// TIA Portal project "Project3" (V13)

(* hardware
DEVICE "S7-1200 station_1"  S7-1200 Station
   slot 0: "Rack_0"  Rack  V1.0
   slot 1: "PLC_1"  CPU 1212C AC/DC/Rly  6ES7 212-1BE40-0XB0  V4.1
DEVICE "GSD device_1"  GSD.Device.PN
   slot 0: "Rack"  Rail  V1.0
   slot 0: "AL1100"  AL1100
   slot 1: "4 Ports_1"  AL1100
DEVICE "HMI_2"  KTP400 Basic PN
   slot 0: "HMI"  HMI  6AV2 123-2DB03-0AX0  13.0.0.0
   slot 1: "HMI_RT_2"  KTP400 Basic PN  6AV2 123-2DB03-0AX0  13.0.0.0
   slot 5: "HMI_2.IE_CP_1"  PROFINET Interface
      slot 1: "PROFINET Interface_1"  PROFINET Interface
         slot 1: "Port_1"  Port
*)

// ===== PLC "PLC_1"  CPU 1212C AC/DC/Rly =====

VAR_GLOBAL   // PLC tag table "Default tag table"
   "Tag_1" AT %Q0.0 : Bool;
   "Tag_2" AT %M0.0 : Bool;
   "System_Byte" AT %MB1 : Byte;
   "FirstScan" AT %M1.0 : Bool;
   "DiagStatusUpdate" AT %M1.1 : Bool;
   "AlwaysTRUE" AT %M1.2 : Bool;
   "AlwaysFALSE" AT %M1.3 : Bool;
   "Clock_Byte" AT %MB0 : Byte;
   "Clock_5Hz" AT %M0.1 : Bool;
   "Clock_2.5Hz" AT %M0.2 : Bool;
   "Clock_2Hz" AT %M0.3 : Bool;
   "Clock_1.25Hz" AT %M0.4 : Bool;
   "Clock_1Hz" AT %M0.5 : Bool;
   "Clock_0.625Hz" AT %M0.6 : Bool;
   "Clock_0.5Hz" AT %M0.7 : Bool;
   "Tag_3" AT %M10.0 : Bool;
END_VAR

VAR_GLOBAL   // PLC tag table "RFID"
   "i_command_value" AT %IB90 : Byte;
   "i_command_ack" AT %I91.0 : Bool;
   "i_command_end" AT %I91.1 : Bool;
   "i_tag_present" AT %I91.2 : Bool;
   "i_antenna_deactivated" AT %I91.3 : Bool;
   "i_read_value_0" AT %IW92 : Int;
   "i_read_value_1" AT %IW94 : Int;
   "i_read_value_2" AT %IW96 : Int;
   "i_read_value_3" AT %IW98 : Int;
   "q_command_value" AT %QB84 : Byte;
   "q_start_r/w" AT %Q85.0 : Bool;
   "q_antenna_deactivate" AT %Q85.3 : Bool;
   "q_write_value_0" AT %QW86 : Int;
   "q_write_value_1" AT %QW88 : Int;
   "q_write_value_2" AT %QW90 : Int;
   "q_write_value_3" AT %QW92 : Int;
END_VAR

TYPE "RFID_IOLink"
   STRUCT
      Input : Struct
      END_STRUCT;
      Output : Struct
      END_STRUCT;
   END_STRUCT;
END_TYPE

DATA_BLOCK "test"   // DB2
{ S7_Optimized_Access := 'FALSE' }
VERSION : 0.1
   VAR
      demo : Bool;
      data : Int;
   END_VAR
BEGIN
END_DATA_BLOCK

DATA_BLOCK "Logic_DB"   // DB4
{ S7_Optimized_Access := 'FALSE' }
VERSION : 0.1
// stored: InstanceOfName Logic
"Logic"
BEGIN
END_DATA_BLOCK

// folder: RFID

DATA_BLOCK "RFIDData"   // DB1
{ S7_Optimized_Access := 'FALSE' }
VERSION : 0.1
   VAR
      RFID : "RFID_IOLink";
   END_VAR
BEGIN
END_DATA_BLOCK

DATA_BLOCK "Logic DB"   // DB3
{ S7_Optimized_Access := 'FALSE' }
VERSION : 0.1
   VAR
      TimeParameters : Struct
      END_STRUCT;
      BufferControl : Struct
      END_STRUCT;
      Error : Struct
      END_STRUCT;
   END_VAR
BEGIN
END_DATA_BLOCK

DATA_BLOCK "BufferData_DB"   // DB5
{ S7_Optimized_Access := 'FALSE' }
VERSION : 0.1
// stored: InstanceOfName BufferData
"BufferData"
BEGIN
END_DATA_BLOCK

// folder: (top level)

ORGANIZATION_BLOCK "Main"   // OB1, LAD, ProgramCycle
TITLE = "Main Program Sweep (Cycle)"
{ S7_Optimized_Access := 'FALSE' }
VERSION : 0.1
BEGIN

REGION Network 1: Read values from RFID
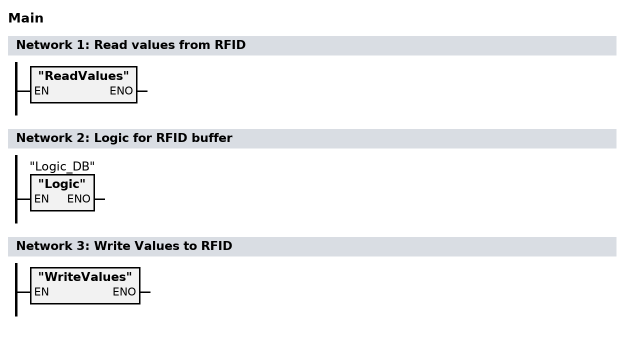
   RUNG wire#powerrail
      "ReadValues"()
   END_RUNG
   // the same network as SCL:
   "ReadValues"();
END_REGION

REGION Network 2: Logic for RFID buffer
   RUNG wire#powerrail
      "Logic_DB"()
   END_RUNG
   // the same network as SCL:
   "Logic_DB"();   // "Logic"
END_REGION

REGION Network 3: Write Values to RFID
   RUNG wire#powerrail
      "WriteValues"()
   END_RUNG
   // the same network as SCL:
   "WriteValues"();
END_REGION
END_ORGANIZATION_BLOCK

// folder: RFID

FUNCTION_BLOCK "Logic"   // FB1, FBD
{ S7_Optimized_Access := 'FALSE' }
VERSION : 0.1
BEGIN

REGION Network 1: Log of tags with timestamp
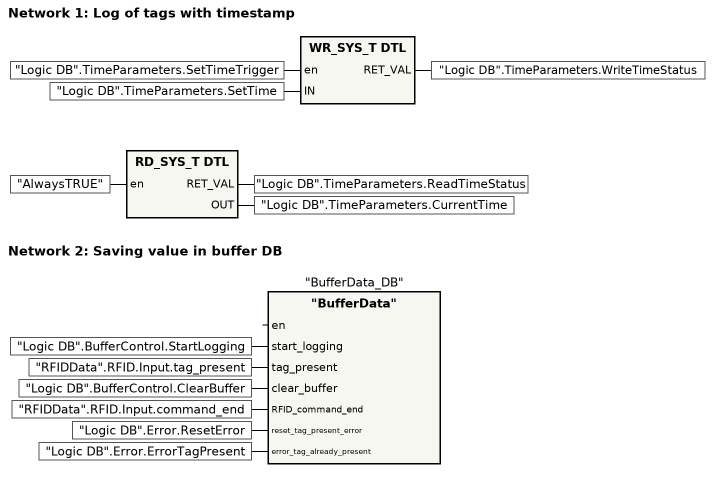
   IF "Logic DB".TimeParameters.SetTimeTrigger THEN
       "Logic DB".TimeParameters.WriteTimeStatus := WR_SYS_T(IN := "Logic DB".TimeParameters.SetTime);
   END_IF;
   IF "AlwaysTRUE" THEN
       "Logic DB".TimeParameters.ReadTimeStatus := RD_SYS_T(OUT => "Logic DB".TimeParameters.CurrentTime);
   END_IF;
END_REGION

REGION Network 2: Saving value in buffer DB
   "BufferData_DB"(start_logging := "Logic DB".BufferControl.StartLogging,   // "BufferData"
                   tag_present := "RFIDData".RFID.Input.tag_present,
                   clear_buffer := "Logic DB".BufferControl.ClearBuffer,
                   RFID_command_end := "RFIDData".RFID.Input.command_end,
                   reset_tag_present_error := "Logic DB".Error.ResetError,
                   error_tag_already_present := "Logic DB".Error.ErrorTagPresent);
END_REGION
END_FUNCTION_BLOCK

FUNCTION_BLOCK "BufferData"   // FB2, SCL
{ S7_Optimized_Access := 'FALSE' }
VERSION : 0.1
BEGIN
   //Generating rising edge bit for RFID 'End' status
   #command_end_flag:= #RFID_command_end AND NOT #M_command_end_flag;
   #M_command_end_flag := #RFID_command_end;

   //Check tag validity i.e. Tag should not be = 0 and not already registered
   IF (#start_logging AND NOT #error_tag_already_present) THEN
       IF (#command_end_flag) AND ("RFIDData".RFID.Input.read_values[0] <> 0) THEN 
           FOR #c := 0 TO 5 DO
               IF ("Logic DB".BufferControl.Job[#c].RFID = "RFIDData".RFID.Input.read_values[0]) THEN
                   #error_tag_already_present := true;
                   GOTO x2;
               END_IF;
           END_FOR;
   //IF RFID tag is not registered --> Registering the tag information in the next available slot
           FOR #d := 0 TO 5 DO
               IF (#command_end_flag) AND ("Logic DB".BufferControl.Job[#d].RFID = 0) AND NOT #error_tag_already_present THEN
                   "Logic DB".BufferControl.Job[#d].Job_ID := #d +1;
                   "Logic DB".BufferControl.Job[#d].RFID := "RFIDData".RFID.Input.read_values[0];
                   "Logic DB".BufferControl.Job[#d].ProcessTime :="Logic DB".TimeParameters.CurrentTime ;
                   GOTO x2;
               END_IF;
           END_FOR;
       x2: ;
      END_IF;
   END_IF;

   //Clear log button
   IF #clear_buffer THEN
       FOR #i := 0 TO 5 DO
           "Logic DB".BufferControl.Job[#i].ProcessTime := "Logic DB".TimeParameters.ResetTime;
           "Logic DB".BufferControl.Job[#i].RFID := 0;
           "Logic DB".BufferControl.Job[#i].Job_ID := 0;
       END_FOR;

   END_IF;

   IF (#reset_tag_present_error) THEN
       #error_tag_already_present := false;
   END_IF;
END_FUNCTION_BLOCK

FUNCTION "ReadValues" : Void   // FC1, SCL
{ S7_Optimized_Access := 'FALSE' }
VERSION : 0.1
BEGIN
   //Reading value from RFID
   "RFIDData".RFID.Input.command_ack:="i_command_ack";
   "RFIDData".RFID.Input.command_value:="i_command_value";
   "RFIDData".RFID.Input.command_end:="i_command_end";
   "RFIDData".RFID.Input.tag_present:="i_tag_present";
   "RFIDData".RFID.Input.Antenna_deactivated:="i_antenna_deactivated";
   "RFIDData".RFID.Input.read_values[0]:="i_read_value_0";
   "RFIDData".RFID.Input.read_values[1]:="i_read_value_1";
   "RFIDData".RFID.Input.read_values[2]:="i_read_value_2";
   "RFIDData".RFID.Input.read_values[3]:="i_read_value_3";
END_FUNCTION

FUNCTION "WriteValues" : Void   // FC2, SCL
{ S7_Optimized_Access := 'FALSE' }
VERSION : 0.1
BEGIN
   //Writing values to RFID
   "q_command_value" := "RFIDData".RFID.Output.command_value;
   "q_start_r/w" := "RFIDData".RFID.Output."Start_r/w";
   "q_antenna_deactivate" := "RFIDData".RFID.Output.Deactivate_antenna;
   "q_write_value_0" := "RFIDData".RFID.Output.write_values[0];
   "q_write_value_1" := "RFIDData".RFID.Output.write_values[1];
   "q_write_value_2" := "RFIDData".RFID.Output.write_values[2];
   "q_write_value_3" := "RFIDData".RFID.Output.write_values[3];
END_FUNCTION

(* ===== HMI "HMI_RT_2" =====
connection "HMI_Connection_1": ETHERNET, SMART_S7_1200_OMS

HMI tags "RFID"
   "i_command_ack" : Bool, 100 ms
   "i_command_end" : Bool, 100 ms
   "i_tag_present" : Bool, 100 ms
   "i_antenna_deactivated" : Bool, 100 ms
   "i_command_value" : Byte, 100 ms
   "i_read_value_0" : Int, 100 ms
   "i_read_value_1" : Int, 100 ms
   "i_read_value_2" : Int, 100 ms
   "i_read_value_3" : Int, 100 ms
   "q_startr/w" : Bool, 100 ms
   "q_deactivate_antenna" : Bool, 100 ms
   "q_command_value" : Byte, 100 ms
   "q_write_values_0" : Int, 100 ms
   "q_write_values_1" : Int, 100 ms
   "q_write_values_2" : Int, 100 ms
   "q_write_values_3" : Int, 100 ms

text list "command_value": 0 ''; 1 ''; 2 ''; 3 ''; 4 ''

Template "Template_1" 480x272
   Button "Template_Button" at 439,242 size 40x29

screen "Read and write" 480x272, template "Template_1"
   TextField "Text field_1" at 13,9 size 161x22
   TextField "Text field_2" at 17,34 size 99x46
   IOField "I/O field_1" at 125,39 size 99x39
   IOField "I/O field_2" at 125,84 size 99x39
   IOField "I/O field_3" at 125,128 size 99x39
   IOField "I/O field_4" at 125,173 size 99x39
   TextField "Text field_7" at 8,224 size 113x22
   TextField "Text field_8" at 6,243 size 108x22
   TextField "Text field_9" at 149,225 size 94x22
   TextField "Text field_10" at 149,244 size 116x22
   TextField "Text field_3" at 17,79 size 99x46
   TextField "Text field_4" at 17,124 size 99x46
   TextField "Text field_5" at 17,170 size 99x46
   Switch "Switch_1" at 298,231 size 132x33
   TextField "Text field_6" at 246,9 size 165x22
   TextField "Text field_11" at 252,34 size 102x46
   IOField "I/O field_5" at 361,39 size 99x39
   IOField "I/O field_6" at 361,84 size 99x39
   IOField "I/O field_7" at 361,128 size 99x39
   IOField "I/O field_8" at 361,173 size 99x39
   TextField "Text field_12" at 252,78 size 102x46
   TextField "Text field_13" at 252,123 size 102x46
   TextField "Text field_14" at 252,168 size 102x46
*)